Fanuc KAREL source: KA00150.KL

PROGRAM KA00150
%NOLOCKGROUP
VAR
  SRC: ARRAY[4] OF INTEGER
  DST: ARRAY[4] OF SHORT
BEGIN
  DST = SRC
END KA00150
